(****************************************************************************************************<br>
© Syntegon Group.<br>
All rights reserved, also regarding any disposal, exploitation, reproduction, editing, distribution,<br>
as well as in the event of applications for industrial property rights.<br>
*****************************************************************************************************<br>
DESCRIPTION:<br>
Housekeeping: drops invalid entries and products that have travelled beyond vi_lr_BeltX (along the<br>
conveyor from its start). Products a robot is working on (ASSIGNED or PICKED) are kept wherever they are.<br>
The entries that stay move up in runs (usually one: the products leaving are the oldest, at the front).<br>
*****************************************************************************************************<br>
OUTPUT VALUES:<br>
Number of removed entries.<br>
****************************************************************************************************)
METHOD m_RemoveProductsBeyond : UINT
VAR_INPUT
	vi_lr_BeltX							: LREAL;	// [mm] e.g. belt length + some margin so missed products stay visible briefly
END_VAR
VAR
	un_TempCount						: UINT;	// [-] entries before
	un_TempRead							: UINT;
	un_TempWrite						: UINT;
	un_TempRunStart						: UINT;	// [-] first entry of a run of entries that stay
	b_TempStays							: BOOL;
END_VAR
m_RemoveProductsBeyond := 0;
un_TempCount := vo_Visu.stState.nProductCount;
IF un_TempCount = 0 THEN
	RETURN;
END_IF

(* Keep the entries that stay, in order, moving each run of them up in one go. *)
un_TempWrite := 0;
un_TempRead := 0;
WHILE un_TempRead < un_TempCount DO
	IF m_StaysInRegister(un_TempRead, vi_lr_BeltX) THEN
		un_TempRunStart := un_TempRead;
		b_TempStays := TRUE;
		WHILE b_TempStays DO
			un_TempRead := un_TempRead + 1;
			b_TempStays := FALSE;
			IF un_TempRead < un_TempCount THEN
				b_TempStays := m_StaysInRegister(un_TempRead, vi_lr_BeltX);
			END_IF
		END_WHILE
		IF un_TempWrite <> un_TempRunStart THEN
			Tc2_System.MEMMOVE(ADR(vo_Visu.stState.aProducts[un_TempWrite]), ADR(vo_Visu.stState.aProducts[un_TempRunStart]),
				UINT_TO_UDINT(un_TempRead - un_TempRunStart) * SIZEOF(ST_VisuProduct));
		END_IF
		un_TempWrite := un_TempWrite + (un_TempRead - un_TempRunStart);
	ELSE
		un_TempRead := un_TempRead + 1;
	END_IF
END_WHILE

(* Invalidate the freed tail. *)
m_RemoveProductsBeyond := un_TempCount - un_TempWrite;
IF un_TempWrite < un_TempCount THEN
	FOR un_TempRead := un_TempWrite TO un_TempCount - 1 DO
		vo_Visu.stState.aProducts[un_TempRead].bValid := FALSE;
	END_FOR
	vo_Visu.stState.nProductCount := un_TempWrite;
	vo_Visu.stState.nTimestamp := m_DcTime();
	b_IndexValid := FALSE;
END_IF
END_METHOD

(****************************************************************************************************<br>
© Syntegon Group.<br>
All rights reserved, also regarding any disposal, exploitation, reproduction, editing, distribution,<br>
as well as in the event of applications for industrial property rights.<br>
*****************************************************************************************************<br>
DESCRIPTION:<br>
The rotation of the conveyor's pose as a row-major 3x3 matrix, R = Rz(fRz) * Ry(fRy) * Rx(fRx) as the contract<br>
defines it (ST_VisuPose) and the visualisation applies it, for m_BeltToMcs and m_McsToBelt.<br>
****************************************************************************************************)
METHOD PRIVATE m_Rotation : BOOL
VAR_OUTPUT
	vo_lr_Rotation						: ARRAY[0..8] OF LREAL;	// [-] row by row
END_VAR
VAR
	lr_TempCx							: LREAL;
	lr_TempSx							: LREAL;
	lr_TempCy							: LREAL;
	lr_TempSy							: LREAL;
	lr_TempCz							: LREAL;
	lr_TempSz							: LREAL;
END_VAR
lr_TempCx := COS(vo_Visu.stConfig.stPose.fRx * VISU_GlobalConst.VISU_lr_DEG_TO_RAD);
lr_TempSx := SIN(vo_Visu.stConfig.stPose.fRx * VISU_GlobalConst.VISU_lr_DEG_TO_RAD);
lr_TempCy := COS(vo_Visu.stConfig.stPose.fRy * VISU_GlobalConst.VISU_lr_DEG_TO_RAD);
lr_TempSy := SIN(vo_Visu.stConfig.stPose.fRy * VISU_GlobalConst.VISU_lr_DEG_TO_RAD);
lr_TempCz := COS(vo_Visu.stConfig.stPose.fRz * VISU_GlobalConst.VISU_lr_DEG_TO_RAD);
lr_TempSz := SIN(vo_Visu.stConfig.stPose.fRz * VISU_GlobalConst.VISU_lr_DEG_TO_RAD);
vo_lr_Rotation[0] := lr_TempCz * lr_TempCy;
vo_lr_Rotation[1] := lr_TempCz * lr_TempSy * lr_TempSx - lr_TempSz * lr_TempCx;
vo_lr_Rotation[2] := lr_TempCz * lr_TempSy * lr_TempCx + lr_TempSz * lr_TempSx;
vo_lr_Rotation[3] := lr_TempSz * lr_TempCy;
vo_lr_Rotation[4] := lr_TempSz * lr_TempSy * lr_TempSx + lr_TempCz * lr_TempCx;
vo_lr_Rotation[5] := lr_TempSz * lr_TempSy * lr_TempCx - lr_TempCz * lr_TempSx;
vo_lr_Rotation[6] := -lr_TempSy;
vo_lr_Rotation[7] := lr_TempCy * lr_TempSx;
vo_lr_Rotation[8] := lr_TempCy * lr_TempCx;
m_Rotation := TRUE;
END_METHOD

(****************************************************************************************************<br>
© Syntegon Group.<br>
All rights reserved, also regarding any disposal, exploitation, reproduction, editing, distribution,<br>
as well as in the event of applications for industrial property rights.<br>
*****************************************************************************************************<br>
DESCRIPTION:<br>
Sets the belt position: how far the belt surface has travelled, continuous (no modulo).<br>
Call once per cycle; it also stamps the state with the cycle's DC time.<br>
****************************************************************************************************)
METHOD m_SetBeltPosition : BOOL
VAR_INPUT
	vi_lr_Position						: LREAL;	// [mm]
END_VAR
vo_Visu.stState.fBeltPosition := vi_lr_Position;
vo_Visu.stState.nTimestamp := m_DcTime();
m_SetBeltPosition := TRUE;
END_METHOD

(****************************************************************************************************<br>
© Syntegon Group.<br>
All rights reserved, also regarding any disposal, exploitation, reproduction, editing, distribution,<br>
as well as in the event of applications for industrial property rights.<br>
*****************************************************************************************************<br>
DESCRIPTION:<br>
Sets whether the belt is drawn as a body. A conveyor without one (FALSE) shows only its products, zones and<br>
its axis from the origin to the conveying direction arrow. Default TRUE. TRUE if anything changed.<br>
****************************************************************************************************)
METHOD m_SetBodyVisible : BOOL
VAR_INPUT
	vi_b_Visible						: BOOL;	// TRUE = drawn as a body, FALSE = a conveyor without one
END_VAR
VAR
	TempNew								: ST_VisuConveyorConfig;
END_VAR
TempNew := vo_Visu.stConfig;
TempNew.bBody := vi_b_Visible;
m_SetBodyVisible := m_ApplyConfig(TempNew);
END_METHOD

(****************************************************************************************************<br>
© Syntegon Group.<br>
All rights reserved, also regarding any disposal, exploitation, reproduction, editing, distribution,<br>
as well as in the event of applications for industrial property rights.<br>
*****************************************************************************************************<br>
DESCRIPTION:<br>
Sets or clears the fault of the conveyor: drawn red with the message while active. The fault stays until it<br>
is cleared with m_SetFault(vi_b_Active := FALSE, vi_str_Message := ''). TRUE.<br>
****************************************************************************************************)
METHOD m_SetFault : BOOL
VAR_INPUT
	vi_b_Active							: BOOL;	// TRUE: fault active
	vi_str_Message						: STRING(80);	// shown to the operator; empty shows 'Fault'
END_VAR
vo_Visu.stState.stFault.bActive := vi_b_Active;
vo_Visu.stState.stFault.sMessage := vi_str_Message;
m_SetFault := TRUE;
END_METHOD

(****************************************************************************************************<br>
© Syntegon Group.<br>
All rights reserved, also regarding any disposal, exploitation, reproduction, editing, distribution,<br>
as well as in the event of applications for industrial property rights.<br>
*****************************************************************************************************<br>
DESCRIPTION:<br>
Like m_SetBeltPosition, for a modulo axis: unwraps the position so the belt position stays continuous.<br>
Call once per cycle.<br>
*****************************************************************************************************<br>
LIMITS:<br>
The axis must move less than half a modulo period per cycle.<br>
****************************************************************************************************)
METHOD m_SetModuloBeltPosition : BOOL
VAR_INPUT
	vi_lr_ModuloPosition				: LREAL;	// [mm] in [0, vi_lr_ModuloPeriod)
	vi_lr_ModuloPeriod					: LREAL;	// [mm] <= 0 passes vi_lr_ModuloPosition through unchanged
	vi_b_Reset							: BOOL;	// TRUE: restart the belt position at vi_lr_ModuloPosition
END_VAR
VAR
	lr_TempPosition						: LREAL;	// [mm]
	lr_TempDelta						: LREAL;	// [mm]
END_VAR
IF vi_b_Reset OR NOT b_ModuloInitialised OR vi_lr_ModuloPeriod <= 0 THEN
	lr_TempPosition := vi_lr_ModuloPosition;
	b_ModuloInitialised := TRUE;
ELSE
	lr_TempDelta := vi_lr_ModuloPosition - lr_LastModuloPosition;
	IF lr_TempDelta > vi_lr_ModuloPeriod / 2 THEN
		lr_TempDelta := lr_TempDelta - vi_lr_ModuloPeriod;
	ELSIF lr_TempDelta < -vi_lr_ModuloPeriod / 2 THEN
		lr_TempDelta := lr_TempDelta + vi_lr_ModuloPeriod;
	END_IF
	lr_TempPosition := vo_Visu.stState.fBeltPosition + lr_TempDelta;
END_IF
lr_LastModuloPosition := vi_lr_ModuloPosition;
m_SetModuloBeltPosition := m_SetBeltPosition(lr_TempPosition);
END_METHOD

(****************************************************************************************************<br>
© Syntegon Group.<br>
All rights reserved, also regarding any disposal, exploitation, reproduction, editing, distribution,<br>
as well as in the event of applications for industrial property rights.<br>
*****************************************************************************************************<br>
DESCRIPTION:<br>
Moves the conveyor's coordinate system away from the belt start (stPose), in the belt's local frame. Belt<br>
coordinates (zones' start, end and CCS offset) then count from the shifted origin. TRUE if anything changed.<br>
****************************************************************************************************)
METHOD m_SetOriginShift : BOOL
VAR_INPUT
	vi_lr_X								: LREAL;	// [mm] along the conveying direction
	vi_lr_Y								: LREAL;	// [mm] across the belt, 0 = none
	vi_lr_Z								: LREAL;	// [mm] along the belt surface normal, 0 = none
END_VAR
VAR
	TempNew								: ST_VisuConveyorConfig;
END_VAR
TempNew := vo_Visu.stConfig;
TempNew.stOriginShift.fX := vi_lr_X;
TempNew.stOriginShift.fY := vi_lr_Y;
TempNew.stOriginShift.fZ := vi_lr_Z;
m_SetOriginShift := m_ApplyConfig(TempNew);
END_METHOD

(****************************************************************************************************<br>
© Syntegon Group.<br>
All rights reserved, also regarding any disposal, exploitation, reproduction, editing, distribution,<br>
as well as in the event of applications for industrial property rights.<br>
*****************************************************************************************************<br>
DESCRIPTION:<br>
Marks a product of the register to single it out, e.g. as a sample: the visualisation draws it in the mark's<br>
colour instead of its state colour. 0 removes the mark. The mark stays through m_SetProductState and<br>
m_MoveProduct; a product latched again (e.g. put down on another conveyor) enters unmarked, so mark it there<br>
again. Name the marks once with _FC_VisuSetMarkName.<br>
*****************************************************************************************************<br>
OUTPUT VALUES:<br>
FALSE if the product is not in the register or vi_un_Mark is above VISU_un_MAX_MARKS.<br>
****************************************************************************************************)
METHOD m_SetProductMark : BOOL
VAR_INPUT
	vi_udn_Id							: UDINT;	// [-] product id
	vi_un_Mark							: UINT;	// [-] product mark 1..VISU_un_MAX_MARKS, 0 = none
END_VAR
VAR
	n_TempIndex							: INT;
END_VAR
m_SetProductMark := FALSE;
IF vi_un_Mark > VISU_GlobalConst.VISU_un_MAX_MARKS THEN
	RETURN;
END_IF
n_TempIndex := m_FindProduct(vi_udn_Id);
IF n_TempIndex < 0 THEN
	RETURN;
END_IF
IF vo_Visu.stState.aProducts[n_TempIndex].nMark <> vi_un_Mark THEN
	vo_Visu.stState.aProducts[n_TempIndex].nMark := vi_un_Mark;
	vo_Visu.stState.nTimestamp := m_DcTime();
END_IF
m_SetProductMark := TRUE;
END_METHOD

(****************************************************************************************************<br>
© Syntegon Group.<br>
All rights reserved, also regarding any disposal, exploitation, reproduction, editing, distribution,<br>
as well as in the event of applications for industrial property rights.<br>
*****************************************************************************************************<br>
DESCRIPTION:<br>
Changes a product's state and names the client that changed it: the robot that is assigned to, picks,<br>
places or releases it, the station that rejects it. The state before is kept as ePreviousState when the<br>
state changes; calling it again with the same state keeps it. The product keeps its mark.<br>
FALSE if the product is not in the register.<br>
****************************************************************************************************)
METHOD m_SetProductState : BOOL
VAR_INPUT
	vi_udn_Id							: UDINT;	// [-] product id
	vi_e_State							: E_VisuProductState;
	vi_udn_ClientId						: UDINT;	// [-] manifest id of the client making the change, 0 = none
	vi_udn_MoverId						: UDINT;	// [-] mover of an XTS gantry or loop carrying the product, 0 = none
	vi_udn_FingerId						: UDINT;	// [-] gripper finger (1-based) the product hangs from while picked, 0 = the flange
END_VAR
VAR
	n_TempIndex							: INT;
END_VAR
n_TempIndex := m_FindProduct(vi_udn_Id);
m_SetProductState := n_TempIndex >= 0;
IF m_SetProductState THEN
	IF vo_Visu.stState.aProducts[n_TempIndex].eState <> vi_e_State THEN
		vo_Visu.stState.aProducts[n_TempIndex].ePreviousState := vo_Visu.stState.aProducts[n_TempIndex].eState;
	END_IF
	vo_Visu.stState.aProducts[n_TempIndex].eState := vi_e_State;
	vo_Visu.stState.aProducts[n_TempIndex].nLastClientId := vi_udn_ClientId;
	vo_Visu.stState.aProducts[n_TempIndex].nMoverId := vi_udn_MoverId;
	vo_Visu.stState.aProducts[n_TempIndex].nFingerId := vi_udn_FingerId;
	vo_Visu.stState.nTimestamp := m_DcTime();
END_IF
END_METHOD

(****************************************************************************************************<br>
© Syntegon Group.<br>
All rights reserved, also regarding any disposal, exploitation, reproduction, editing, distribution,<br>
as well as in the event of applications for industrial property rights.<br>
*****************************************************************************************************<br>
DESCRIPTION:<br>
Adds a product type, or updates the one with the same id. FALSE for vi_udn_Id = 0 or a full list. A CYLINDER's<br>
length and width are its diameters (equal: round, different: oval).<br>
****************************************************************************************************)
METHOD m_SetProductType : BOOL
VAR_INPUT
	vi_udn_Id							: UDINT;	// [-] referenced by m_LatchProduct's vi_udn_ProductType
	vi_lr_Length						: LREAL;	// [mm] along the conveying direction
	vi_lr_Width							: LREAL;	// [mm]
	vi_lr_Height						: LREAL;	// [mm]
	vi_e_Shape							: E_VisuProductShape;	// [-] solid of the product, BOX for a plain box
	vi_lr_CornerRadius					: LREAL;	// [mm] rounded vertical edges of a ROUNDED_BOX, 0 for other shapes
END_VAR
VAR
	TempNew								: ST_VisuConveyorConfig;
	un_TempIndex						: UINT;
END_VAR
m_SetProductType := FALSE;
IF vi_udn_Id = 0 THEN
	RETURN;
END_IF
TempNew := vo_Visu.stConfig;
un_TempIndex := 0;
(* ST evaluates both operands of AND: test the index before reading the array. *)
WHILE un_TempIndex < TempNew.nProductTypeCount DO
	IF TempNew.aProductTypes[un_TempIndex].nId = vi_udn_Id THEN
		EXIT;
	END_IF
	un_TempIndex := un_TempIndex + 1;
END_WHILE
IF un_TempIndex >= VISU_GlobalConst_Param.VISU_un_MAX_PRODUCT_TYPES THEN
	RETURN;
END_IF
IF un_TempIndex = TempNew.nProductTypeCount THEN
	TempNew.nProductTypeCount := TempNew.nProductTypeCount + 1;
END_IF
TempNew.aProductTypes[un_TempIndex].nId := vi_udn_Id;
TempNew.aProductTypes[un_TempIndex].fLength := vi_lr_Length;
TempNew.aProductTypes[un_TempIndex].fWidth := vi_lr_Width;
TempNew.aProductTypes[un_TempIndex].fHeight := vi_lr_Height;
TempNew.aProductTypes[un_TempIndex].eShape := vi_e_Shape;
TempNew.aProductTypes[un_TempIndex].fCornerRadius := vi_lr_CornerRadius;
m_ApplyConfig(TempNew);
m_SetProductType := TRUE;
END_METHOD

(****************************************************************************************************<br>
© Syntegon Group.<br>
All rights reserved, also regarding any disposal, exploitation, reproduction, editing, distribution,<br>
as well as in the event of applications for industrial property rights.<br>
*****************************************************************************************************<br>
DESCRIPTION:<br>
Whether register entry vi_un_Index stays in the register for m_RemoveProductsBeyond: it is valid and has not<br>
travelled beyond vi_lr_BeltX, or a robot is working on it (ASSIGNED or PICKED).<br>
****************************************************************************************************)
METHOD PRIVATE m_StaysInRegister : BOOL
VAR_INPUT
	vi_un_Index							: UINT;	// [-] register index
	vi_lr_BeltX							: LREAL;	// [mm] along the conveyor from its start
END_VAR
(* Belt X from the belt start: the latch pose counts from the origin shift and moves with the belt travel. *)
m_StaysInRegister := vo_Visu.stState.aProducts[vi_un_Index].bValid
	AND (vo_Visu.stConfig.stOriginShift.fX + vo_Visu.stState.aProducts[vi_un_Index].stLatchPose.fX
			+ vo_Visu.stState.fBeltPosition - vo_Visu.stState.aProducts[vi_un_Index].fLatchBeltPosition <= vi_lr_BeltX
		OR vo_Visu.stState.aProducts[vi_un_Index].eState = E_VisuProductState.ASSIGNED
		OR vo_Visu.stState.aProducts[vi_un_Index].eState = E_VisuProductState.PICKED);
END_METHOD

END_FUNCTION_BLOCK

// POUs/_FB_VisuComponent
(****************************************************************************************************<br>
© Syntegon Group.<br>
All rights reserved, also regarding any disposal, exploitation, reproduction, editing, distribution,<br>
as well as in the event of applications for industrial property rights.<br>
*****************************************************************************************************<br>
DESCRIPTION:<br>
Base of every visualised component (_FB_VisuConveyor, _FB_VisuDelta, ...). Handles the manifest entry,<br>
the config version and the DC timestamps. Not used directly.<br>
*****************************************************************************************************<br>
VERSION         ¦ DATE       ¦ NAME      ¦ CHANGE<br>
Syn_Visu 3.0.0  ¦ 2026-10-31 ¦ J.Willner ¦ Naming and layout after the TCAT programming guideline<br>
Syn_Visu 8.0.0  ¦ 2026-11-05 ¦ J.Willner ¦ m_Register without vi_str_Path: the symbol path comes from the instance path<br>
Syn_Visu 10.0.0 ¦ 2026-11-14 ¦ J.Willner ¦ m_SetPose for every component; symbol path from _FC_VisuSymbolPath<br>
****************************************************************************************************)
{attribute 'reflection'}
FUNCTION_BLOCK ABSTRACT _FB_VisuComponent
VAR
	RefManifest							: REFERENCE TO ST_VisuManifest;	// set by m_Register
	udn_ComponentId						: UDINT;	// [-] manifest id, 0 = not registered
	(* Device tree path of this instance, e.g. 'RPP_Visu.Syn_Visu_Demo.MAIN.fb_Infeed', set by TwinCAT at initialisation. *)
	{attribute 'instance-path'}
	{attribute 'noinit'}
	str_InstancePath					: STRING(255);
	str_SymbolPath						: STRING(255);	// symbol path of vo_Visu for the manifest, from str_InstancePath on the first m_Register
END_VAR

(****************************************************************************************************<br>
© Syntegon Group.<br>
All rights reserved, also regarding any disposal, exploitation, reproduction, editing, distribution,<br>
as well as in the event of applications for industrial property rights.<br>
*****************************************************************************************************<br>
DESCRIPTION:<br>
Manifest type of the component. Overridden by every derived FB.<br>
****************************************************************************************************)
METHOD PROTECTED m_ComponentType : E_VisuComponentType
m_ComponentType := E_VisuComponentType.NONE;
END_METHOD

(****************************************************************************************************<br>
© Syntegon Group.<br>
All rights reserved, also regarding any disposal, exploitation, reproduction, editing, distribution,<br>
as well as in the event of applications for industrial property rights.<br>
*****************************************************************************************************<br>
DESCRIPTION:<br>
Distributed-clock time of the calling task's current cycle in ns since 2000-01-01; 0 if unknown.<br>
****************************************************************************************************)
METHOD PROTECTED m_DcTime : ULINT
VAR
	dn_TempTaskIndex					: DINT;
END_VAR
dn_TempTaskIndex := Tc2_System.GETCURTASKINDEXEX();
IF dn_TempTaskIndex > 0 THEN
	m_DcTime := LINT_TO_ULINT(TwinCAT_SystemInfoVarList._TaskInfo[dn_TempTaskIndex].DcTaskTime);
ELSE
	m_DcTime := 0;
END_IF
END_METHOD

(****************************************************************************************************<br>
© Syntegon Group.<br>
All rights reserved, also regarding any disposal, exploitation, reproduction, editing, distribution,<br>
as well as in the event of applications for industrial property rights.<br>
*****************************************************************************************************<br>
DESCRIPTION:<br>
Manifest id given to m_Register; 0 while not registered.<br>
****************************************************************************************************)
METHOD m_Id : UDINT
m_Id := udn_ComponentId;
END_METHOD

(****************************************************************************************************<br>
© Syntegon Group.<br>
All rights reserved, also regarding any disposal, exploitation, reproduction, editing, distribution,<br>
as well as in the event of applications for industrial property rights.<br>
*****************************************************************************************************<br>
DESCRIPTION:<br>
Increments the manifest's nConfigVersion so the gateway re-reads the config. No effect before m_Register.<br>
****************************************************************************************************)
METHOD PROTECTED m_NotifyConfigChanged : BOOL
m_NotifyConfigChanged := __ISVALIDREF(RefManifest);
IF m_NotifyConfigChanged THEN
	RefManifest.nConfigVersion := RefManifest.nConfigVersion + 1;
END_IF
END_METHOD

(****************************************************************************************************<br>
© Syntegon Group.<br>
All rights reserved, also regarding any disposal, exploitation, reproduction, editing, distribution,<br>
as well as in the event of applications for industrial property rights.<br>
*****************************************************************************************************<br>
DESCRIPTION:<br>
Where the derived FB keeps its pose in its contract structure, for m_SetPose.<br>
****************************************************************************************************)
METHOD PROTECTED ABSTRACT m_Pose : BOOL
VAR_OUTPUT
	vo_p_Pose							: POINTER TO ST_VisuPose;
END_VAR
END_METHOD

(****************************************************************************************************<br>
© Syntegon Group.<br>
All rights reserved, also regarding any disposal, exploitation, reproduction, editing, distribution,<br>
as well as in the event of applications for industrial property rights.<br>
*****************************************************************************************************<br>
DESCRIPTION:<br>
Adds this component to the manifest; increments nConfigVersion when the entry is new.<br>
Idempotent: call it every cycle, which also keeps the manifest reference valid after an online change.<br>
The symbol path the gateway reads comes from the instance's own path (see _FC_VisuSymbolPath and<br>
VISU_un_INSTANCE_PATH_SKIP).<br>
*****************************************************************************************************<br>
OUTPUT VALUES:<br>
FALSE for vi_udn_Id = 0, an id already used by a different entry, or a full manifest.<br>
****************************************************************************************************)
METHOD m_Register : BOOL
VAR_IN_OUT
	vio_Manifest						: ST_VisuManifest;	// GVL_Visu.stManifest of the application
END_VAR
VAR_INPUT
	vi_udn_Id							: UDINT;	// [-] unique, > 0
	vi_str_Name							: STRING(80);	// display name
END_VAR
VAR
	e_TempType							: E_VisuComponentType;
	un_TempIndex						: UINT;
END_VAR
m_Register := FALSE;
RefManifest REF= vio_Manifest;
(* Always report the contract version of the library actually running, also after an online change. *)
vio_Manifest.nProtocolVersion := VISU_GlobalConst.VISU_un_PROTOCOL_VERSION;
vio_Manifest.sLibraryVersion := VISU_GlobalConst.VISU_str_LIBRARY_VERSION;
e_TempType := m_ComponentType();
IF vi_udn_Id = 0 OR e_TempType = E_VisuComponentType.NONE THEN
	RETURN;
END_IF
IF str_SymbolPath = '' THEN
	str_SymbolPath := _FC_VisuSymbolPath(vio_str_InstancePath := str_InstancePath, vi_str_Member := '.vo_Visu');
END_IF

(* An existing entry with the same id must match exactly. *)
un_TempIndex := 0;
WHILE un_TempIndex < vio_Manifest.nCount AND un_TempIndex < VISU_GlobalConst_Param.VISU_un_MAX_MANIFEST_ENTRIES DO
	IF vio_Manifest.aEntries[un_TempIndex].nId = vi_udn_Id THEN
		m_Register := vio_Manifest.aEntries[un_TempIndex].eType = e_TempType
					AND vio_Manifest.aEntries[un_TempIndex].sName = vi_str_Name
					AND vio_Manifest.aEntries[un_TempIndex].sPath = str_SymbolPath;
		IF m_Register THEN
			udn_ComponentId := vi_udn_Id;
		END_IF
		RETURN;
	END_IF
	un_TempIndex := un_TempIndex + 1;
END_WHILE

(* New entry. *)
IF vio_Manifest.nCount >= VISU_GlobalConst_Param.VISU_un_MAX_MANIFEST_ENTRIES THEN
	RETURN;
END_IF
vio_Manifest.aEntries[vio_Manifest.nCount].nId := vi_udn_Id;
vio_Manifest.aEntries[vio_Manifest.nCount].eType := e_TempType;
vio_Manifest.aEntries[vio_Manifest.nCount].sName := vi_str_Name;
vio_Manifest.aEntries[vio_Manifest.nCount].sPath := str_SymbolPath;
vio_Manifest.nCount := vio_Manifest.nCount + 1;
vio_Manifest.nConfigVersion := vio_Manifest.nConfigVersion + 1;
udn_ComponentId := vi_udn_Id;
m_Register := TRUE;
END_METHOD

(****************************************************************************************************<br>
© Syntegon Group.<br>
All rights reserved, also regarding any disposal, exploitation, reproduction, editing, distribution,<br>
as well as in the event of applications for industrial property rights.<br>
*****************************************************************************************************<br>
DESCRIPTION:<br>
Sets the component's pose in the MCS; where it lies on the component (a conveyor's belt start, a Delta's base<br>
centre, ...) says the guide. A parameter FB of Syn_Config sets it with m_PassOn; m_Configure holds only the<br>
hardware. Increments the config version only when the pose changes, so it may be called every cycle.<br>
*****************************************************************************************************<br>
OUTPUT VALUES:<br>
TRUE if the pose changed.<br>
****************************************************************************************************)
METHOD m_SetPose : BOOL
VAR_INPUT
	vi_Pose								: ST_VisuPose;	// MCS
END_VAR
VAR
	p_TempPose							: POINTER TO ST_VisuPose;
END_VAR
m_SetPose := FALSE;
m_Pose(vo_p_Pose => p_TempPose);
IF p_TempPose = 0 THEN
	RETURN;
END_IF
(* ST_VisuPose holds LREALs only, so a memory compare sees no padding. *)
m_SetPose := Tc2_System.MEMCMP(ADR(vi_Pose), p_TempPose, SIZEOF(vi_Pose)) <> 0;
IF m_SetPose THEN
	p_TempPose^ := vi_Pose;
	m_NotifyConfigChanged();
END_IF
END_METHOD

END_FUNCTION_BLOCK

// POUs/_FB_VisuDelta
(****************************************************************************************************<br>
© Syntegon Group.<br>
All rights reserved, also regarding any disposal, exploitation, reproduction, editing, distribution,<br>
as well as in the event of applications for industrial property rights.<br>
*****************************************************************************************************<br>
DESCRIPTION:<br>
One visualised Delta robot. Typical cycle:<br>
  fb_Delta.m_Register(vio_Manifest := GVL_Visu.stManifest, vi_udn_Id := 10, vi_str_Name := 'Delta 1');<br>
  fb_Delta.m_SetPose(vi_Pose := BasePose);<br>
  fb_Delta.m_Configure(vi_lr_BaseRadius := 200, vi_lr_EffectorRadius := 50,<br>
      vi_lr_UpperArmLength := 400, vi_lr_LowerArmLength := 1000);<br>
  fb_Delta.m_SetFinger(vi_un_Finger := 1, vi_lr_Diameter := 40, vi_lr_Height := 50);<br>
  fb_Delta.m_SetWorkingArea(vi_lr_Radius := 750, vi_lr_ZMin := -1300, vi_lr_ZMax := -700, vi_lr_ConeHeight := 200,<br>
      vi_lr_ConeBottomRadius := 450);<br>
  fb_Delta.m_SetLimitArea(vi_lr_XMin := -500, vi_lr_XMax := 500, vi_lr_YMin := -750, vi_lr_YMax := 750,<br>
      vi_lr_ZMin := -1500, vi_lr_ZMax := -700);<br>
  fb_Delta.m_SetZone(vi_un_Zone := 1, vi_udn_ConveyorId := 1, vi_lr_Start := 1100, vi_lr_End := 1900,<br>
      vi_lr_AllocationOffset := 300, vi_lr_CcsOffset := 1100, vi_lr_StartY := 0, vi_lr_EndY := 0);<br>
  fb_Delta.m_SetTcp(vi_ActualTcp := ActualTcp, vi_SetpointTcp := SetpointTcp);<br>
  fb_Delta.m_SetFingerState(vi_un_Finger := 1, vi_Pose := CupPose, vi_b_Active := b_Vacuum);<br>
Only the TCP (the gripper flange) is reported; the visualisation derives the arms from it. Tool rotations<br>
(e.g. a 4th axis) show only through the finger poses, absolute in the MCS. The config methods may be called<br>
every cycle; the config version only changes when a value does.<br>
*****************************************************************************************************<br>
OUTPUT VALUES:<br>
vo_Visu is the contract structure the gateway reads at the path given to m_Register. Do not write it.<br>
*****************************************************************************************************<br>
VERSION         ¦ DATE       ¦ NAME      ¦ CHANGE<br>
Syn_Visu 3.0.0  ¦ 2026-10-31 ¦ J.Willner ¦ Naming and layout after the TCAT programming guideline<br>
Syn_Visu 4.0.0  ¦ 2026-11-01 ¦ J.Willner ¦ Zones and fingers from _FB_VisuRobot; m_SetZone by index, no kind<br>
Syn_Visu 10.0.0 ¦ 2026-11-14 ¦ J.Willner ¦ Pose by m_SetPose, not m_Configure<br>
****************************************************************************************************)
FUNCTION_BLOCK _FB_VisuDelta EXTENDS _FB_VisuRobot
VAR_OUTPUT
	vo_Visu								: ST_VisuDelta;	// contract structure read by the gateway
END_VAR

(****************************************************************************************************<br>
© Syntegon Group.<br>
All rights reserved, also regarding any disposal, exploitation, reproduction, editing, distribution,<br>
as well as in the event of applications for industrial property rights.<br>
*****************************************************************************************************<br>
DESCRIPTION:<br>
Takes over vio_New and increments the config version if it differs from the current config. TRUE if changed.<br>
****************************************************************************************************)
METHOD PRIVATE m_ApplyConfig : BOOL
VAR_IN_OUT
	vio_New								: ST_VisuDeltaConfig;
END_VAR
m_ApplyConfig := Tc2_System.MEMCMP(ADR(vio_New), ADR(vo_Visu.stConfig), SIZEOF(vio_New)) <> 0;
IF m_ApplyConfig THEN
	vo_Visu.stConfig := vio_New;
	m_NotifyConfigChanged();
END_IF
END_METHOD

(****************************************************************************************************<br>
© Syntegon Group.<br>
All rights reserved, also regarding any disposal, exploitation, reproduction, editing, distribution,<br>
as well as in the event of applications for industrial property rights.<br>
*****************************************************************************************************<br>
DESCRIPTION:<br>
Base pose last set by m_SetPose, MCS.<br>
****************************************************************************************************)
METHOD m_BasePose : ST_VisuPose
m_BasePose := vo_Visu.stConfig.stPose;
END_METHOD

(****************************************************************************************************<br>
© Syntegon Group.<br>
All rights reserved, also regarding any disposal, exploitation, reproduction, editing, distribution,<br>
as well as in the event of applications for industrial property rights.<br>
*****************************************************************************************************<br>
DESCRIPTION:<br>
Manifest type: Delta robot.<br>
****************************************************************************************************)
METHOD PROTECTED m_ComponentType : E_VisuComponentType
m_ComponentType := E_VisuComponentType.DELTA;
END_METHOD

(****************************************************************************************************<br>
© Syntegon Group.<br>
All rights reserved, also regarding any disposal, exploitation, reproduction, editing, distribution,<br>
as well as in the event of applications for industrial property rights.<br>
*****************************************************************************************************<br>
DESCRIPTION:<br>
Sets the geometry; its pose (m_SetPose) is the base centre. Arm 1 lies along the base's local +X; arms 2 and 3 follow<br>
counter-clockwise (seen from above) at 120 deg each. TRUE if anything changed.<br>
****************************************************************************************************)
METHOD m_Configure : BOOL
VAR_INPUT
	vi_lr_BaseRadius					: LREAL;	// [mm] base centre to shoulder joint
	vi_lr_EffectorRadius				: LREAL;	// [mm] effector centre to lower-arm joint
	vi_lr_UpperArmLength				: LREAL;	// [mm]
	vi_lr_LowerArmLength				: LREAL;	// [mm]
END_VAR
VAR
	TempNew								: ST_VisuDeltaConfig;
END_VAR
TempNew := vo_Visu.stConfig;
TempNew.fBaseRadius := vi_lr_BaseRadius;
TempNew.fEffectorRadius := vi_lr_EffectorRadius;
TempNew.fUpperArmLength := vi_lr_UpperArmLength;
TempNew.fLowerArmLength := vi_lr_LowerArmLength;
m_Configure := m_ApplyConfig(TempNew);
END_METHOD

(****************************************************************************************************<br>
© Syntegon Group.<br>
All rights reserved, also regarding any disposal, exploitation, reproduction, editing, distribution,<br>
as well as in the event of applications for industrial property rights.<br>
*****************************************************************************************************<br>
DESCRIPTION:<br>
The robot's gripper fingers for _FB_VisuRobot.m_SetFinger and m_ClearFingers.<br>
****************************************************************************************************)
METHOD PROTECTED m_Fingers : BOOL
VAR_OUTPUT
	vo_p_Count							: POINTER TO UINT;
	vo_p_Fingers						: POINTER TO ARRAY[0..VISU_GlobalConst_Param.VISU_un_MAX_FINGERS - 1] OF ST_VisuFinger;
END_VAR
vo_p_Count := ADR(vo_Visu.stConfig.nFingerCount);
vo_p_Fingers := ADR(vo_Visu.stConfig.aFingers);
m_Fingers := TRUE;
END_METHOD

(****************************************************************************************************<br>
© Syntegon Group.<br>
All rights reserved, also regarding any disposal, exploitation, reproduction, editing, distribution,<br>
as well as in the event of applications for industrial property rights.<br>
*****************************************************************************************************<br>
DESCRIPTION:<br>
The robot's limit area and TCP limit area for _FB_VisuRobot.m_SetLimitArea, m_ClearLimitArea,<br>
m_SetTcpLimitArea and m_ClearTcpLimitArea.<br>
****************************************************************************************************)
METHOD PROTECTED m_LimitArea : BOOL
VAR_OUTPUT
	vo_p_LimitArea						: POINTER TO ST_VisuLimitArea;
	vo_p_TcpLimitArea					: POINTER TO ST_VisuLimitArea;
END_VAR
vo_p_LimitArea := ADR(vo_Visu.stConfig.stLimitArea);
vo_p_TcpLimitArea := ADR(vo_Visu.stConfig.stTcpLimitArea);
m_LimitArea := TRUE;
END_METHOD

(****************************************************************************************************<br>
© Syntegon Group.<br>
All rights reserved, also regarding any disposal, exploitation, reproduction, editing, distribution,<br>
as well as in the event of applications for industrial property rights.<br>
*****************************************************************************************************<br>
DESCRIPTION:<br>
The pose in vo_Visu, for m_SetPose.<br>
****************************************************************************************************)
METHOD PROTECTED m_Pose : BOOL
VAR_OUTPUT
	vo_p_Pose							: POINTER TO ST_VisuPose;
END_VAR
vo_p_Pose := ADR(vo_Visu.stConfig.stPose);
m_Pose := TRUE;
END_METHOD

(****************************************************************************************************<br>
© Syntegon Group.<br>
All rights reserved, also regarding any disposal, exploitation, reproduction, editing, distribution,<br>
as well as in the event of applications for industrial property rights.<br>
*****************************************************************************************************<br>
DESCRIPTION:<br>
Sets or clears the fault of the robot: drawn red with the message while active. The fault stays until it<br>
is cleared with m_SetFault(vi_b_Active := FALSE, vi_str_Message := ''). TRUE.<br>
****************************************************************************************************)
METHOD m_SetFault : BOOL
VAR_INPUT
	vi_b_Active							: BOOL;	// TRUE: fault active
	vi_str_Message						: STRING(80);	// shown to the operator; empty shows 'Fault'
END_VAR
vo_Visu.stState.stFault.bActive := vi_b_Active;
vo_Visu.stState.stFault.sMessage := vi_str_Message;
m_SetFault := TRUE;
END_METHOD

(****************************************************************************************************<br>
© Syntegon Group.<br>
All rights reserved, also regarding any disposal, exploitation, reproduction, editing, distribution,<br>
as well as in the event of applications for industrial property rights.<br>
*****************************************************************************************************<br>
DESCRIPTION:<br>
Reports finger vi_un_Finger (1-based): the pose of its frame (centre of its top face), absolute in the MCS,<br>
and whether it grips. Call once per cycle per configured finger. A finger never reported here is drawn at its<br>
offset on the flange (m_SetFingerOffset, ADR 0018).<br>
*****************************************************************************************************<br>
OUTPUT VALUES:<br>
FALSE outside 1..VISU_GlobalConst_Param.VISU_un_MAX_FINGERS.<br>
****************************************************************************************************)
METHOD m_SetFingerState : BOOL
VAR_INPUT
	vi_un_Finger						: UINT;	// [-] 1-based
	vi_Pose								: ST_VisuPose;	// MCS
	vi_b_Active							: BOOL;	// TRUE while the finger grips
END_VAR
m_SetFingerState := vi_un_Finger > 0 AND vi_un_Finger <= VISU_GlobalConst_Param.VISU_un_MAX_FINGERS;
IF m_SetFingerState THEN
	vo_Visu.stState.aFingerStates[vi_un_Finger - 1].stPose := vi_Pose;
	vo_Visu.stState.aFingerStates[vi_un_Finger - 1].bActive := vi_b_Active;
	vo_Visu.stState.aFingerStates[vi_un_Finger - 1].bPoseReported := TRUE;
END_IF
END_METHOD

(****************************************************************************************************<br>
© Syntegon Group.<br>
All rights reserved, also regarding any disposal, exploitation, reproduction, editing, distribution,<br>
as well as in the event of applications for industrial property rights.<br>
*****************************************************************************************************<br>
DESCRIPTION:<br>
Moves the robot's shown coordinate system (origin triad, local measuring coordinates) away from the base<br>
centre (stPose), in the base's local frame. Geometry, working area and limit area stay relative to stPose.<br>
TRUE if anything changed.<br>
****************************************************************************************************)
METHOD m_SetOriginShift : BOOL
VAR_INPUT
	vi_lr_X								: LREAL;	// [mm] along the base's local X
	vi_lr_Y								: LREAL;	// [mm] along the base's local Y, 0 = none
	vi_lr_Z								: LREAL;	// [mm] along the base's local Z, 0 = none
END_VAR
VAR
	TempNew								: ST_VisuDeltaConfig;
END_VAR
TempNew := vo_Visu.stConfig;
TempNew.stOriginShift.fX := vi_lr_X;
TempNew.stOriginShift.fY := vi_lr_Y;
TempNew.stOriginShift.fZ := vi_lr_Z;
m_SetOriginShift := m_ApplyConfig(TempNew);
END_METHOD

(****************************************************************************************************<br>
© Syntegon Group.<br>
All rights reserved, also regarding any disposal, exploitation, reproduction, editing, distribution,<br>
as well as in the event of applications for industrial property rights.<br>
*****************************************************************************************************<br>
DESCRIPTION:<br>
Reports the robot's TCP. Call once per cycle; it also stamps the state with the cycle's DC time.<br>
****************************************************************************************************)
METHOD m_SetTcp : BOOL
VAR_INPUT
	vi_ActualTcp						: ST_VisuPosition;	// MCS, effector centre (the gripper flange)
	vi_SetpointTcp						: ST_VisuPosition;	// MCS
END_VAR
vo_Visu.stState.stActualTcp := vi_ActualTcp;
vo_Visu.stState.stSetpointTcp := vi_SetpointTcp;
vo_Visu.stState.nTimestamp := m_DcTime();
m_SetTcp := TRUE;
END_METHOD

(****************************************************************************************************<br>
© Syntegon Group.<br>
All rights reserved, also regarding any disposal, exploitation, reproduction, editing, distribution,<br>
as well as in the event of applications for industrial property rights.<br>
*****************************************************************************************************<br>
DESCRIPTION:<br>
Sets the working area: a vertical cylinder in the robot frame with an optional cone below. TRUE if changed.<br>
****************************************************************************************************)
METHOD m_SetWorkingArea : BOOL
VAR_INPUT
	vi_lr_Radius						: LREAL;	// [mm]
	vi_lr_ZMin							: LREAL;	// [mm] relative to the base (below the base: negative)
	vi_lr_ZMax							: LREAL;	// [mm] relative to the base
	vi_lr_ConeHeight					: LREAL;	// [mm] below vi_lr_ZMin; 0 = no cone
	vi_lr_ConeBottomRadius				: LREAL;	// [mm]
END_VAR
VAR
	TempNew								: ST_VisuDeltaConfig;
END_VAR
TempNew := vo_Visu.stConfig;
TempNew.stWorkingArea.fRadius := vi_lr_Radius;
TempNew.stWorkingArea.fZMin := vi_lr_ZMin;
TempNew.stWorkingArea.fZMax := vi_lr_ZMax;
TempNew.stWorkingArea.fConeHeight := vi_lr_ConeHeight;
TempNew.stWorkingArea.fConeBottomRadius := vi_lr_ConeBottomRadius;
m_SetWorkingArea := m_ApplyConfig(TempNew);
END_METHOD

(****************************************************************************************************<br>
© Syntegon Group.<br>
All rights reserved, also regarding any disposal, exploitation, reproduction, editing, distribution,<br>
as well as in the event of applications for industrial property rights.<br>
*****************************************************************************************************<br>
DESCRIPTION:<br>
The robot's zones for _FB_VisuZoneComponent.m_SetZone and m_ClearZones.<br>
****************************************************************************************************)
METHOD PROTECTED m_Zones : BOOL
VAR_OUTPUT
	vo_p_Count							: POINTER TO UINT;
	vo_p_Zones							: POINTER TO ARRAY[0..VISU_GlobalConst_Param.VISU_un_MAX_ZONES - 1] OF ST_VisuZone;
END_VAR
vo_p_Count := ADR(vo_Visu.stConfig.nZoneCount);
vo_p_Zones := ADR(vo_Visu.stConfig.aZones);
m_Zones := TRUE;
END_METHOD

END_FUNCTION_BLOCK

// POUs/_FB_VisuRobot
(****************************************************************************************************<br>
© Syntegon Group.<br>
All rights reserved, also regarding any disposal, exploitation, reproduction, editing, distribution,<br>
as well as in the event of applications for industrial property rights.<br>
*****************************************************************************************************<br>
DESCRIPTION:<br>
Base of every robot (Delta, XTS gantry, XTS loop, Cartesian): zones plus the gripper fingers, m_SetFinger,<br>
m_SetFingerOffset (a finger's place on the flange) and m_ClearFingers, the limit area, m_SetLimitArea and<br>
m_ClearLimitArea, and the TCP limit area, m_SetTcpLimitArea and m_ClearTcpLimitArea. A derived FB tells where<br>
its fingers and its boxes lie through m_Fingers and m_LimitArea; an XTS loop has neither box.<br>
Not used directly.<br>
*****************************************************************************************************<br>
VERSION         ¦ DATE       ¦ NAME      ¦ CHANGE<br>
Syn_Visu 4.0.0  ¦ 2026-11-01 ¦ J.Willner ¦ New: fingers shared by all robots<br>
Syn_Visu 9.3.0  ¦ 2026-11-07 ¦ J.Willner ¦ Limit area shared by Delta, XTS gantry and Cartesian (was Delta only)<br>
Syn_Visu 9.4.0  ¦ 2026-11-09 ¦ J.Willner ¦ TCP limit area: m_SetTcpLimitArea, m_ClearTcpLimitArea<br>
Syn_Visu 9.4.1  ¦ 2026-11-09 ¦ J.Willner ¦ Limit area compares ignore padding: no config change from unchanged values<br>
Syn_Visu 9.5.0  ¦ 2026-11-11 ¦ J.Willner ¦ m_SetFingerOffset: a finger's place on the flange (ADR 0018)<br>
****************************************************************************************************)
FUNCTION_BLOCK ABSTRACT _FB_VisuRobot EXTENDS _FB_VisuZoneComponent

(****************************************************************************************************<br>
© Syntegon Group.<br>
All rights reserved, also regarding any disposal, exploitation, reproduction, editing, distribution,<br>
as well as in the event of applications for industrial property rights.<br>
*****************************************************************************************************<br>
DESCRIPTION:<br>
Removes the gripper definition. TRUE if there was one.<br>
****************************************************************************************************)
METHOD m_ClearFingers : BOOL
VAR
	p_TempCount							: POINTER TO UINT;
	p_TempFingers						: POINTER TO ARRAY[0..VISU_GlobalConst_Param.VISU_un_MAX_FINGERS - 1] OF ST_VisuFinger;
	TempEmpty							: ST_VisuFinger;
	un_TempIndex						: UINT;
END_VAR
m_ClearFingers := FALSE;
m_Fingers(vo_p_Count => p_TempCount, vo_p_Fingers => p_TempFingers);
IF p_TempCount = 0 OR p_TempFingers = 0 THEN
	RETURN;
END_IF
m_ClearFingers := p_TempCount^ > 0;
FOR un_TempIndex := 0 TO VISU_GlobalConst_Param.VISU_un_MAX_FINGERS - 1 DO
	p_TempFingers^[un_TempIndex] := TempEmpty;
END_FOR
p_TempCount^ := 0;
IF m_ClearFingers THEN
	m_NotifyConfigChanged();
END_IF
END_METHOD

(****************************************************************************************************<br>
© Syntegon Group.<br>
All rights reserved, also regarding any disposal, exploitation, reproduction, editing, distribution,<br>
as well as in the event of applications for industrial property rights.<br>
*****************************************************************************************************<br>
DESCRIPTION:<br>
Removes the limit area. TRUE if there was one.<br>
****************************************************************************************************)
METHOD m_ClearLimitArea : BOOL
VAR
	p_TempLimitArea						: POINTER TO ST_VisuLimitArea;
	TempEmpty							: ST_VisuLimitArea;
END_VAR
m_ClearLimitArea := FALSE;
m_LimitArea(vo_p_LimitArea => p_TempLimitArea);
IF p_TempLimitArea = 0 THEN
	RETURN;
END_IF
m_ClearLimitArea := p_TempLimitArea^.bActive;
(* Zeroed first: the MEMCMP below also compares the padding after bActive, which a method local leaves undefined. *)
Tc2_System.MEMSET(ADR(TempEmpty), 0, SIZEOF(TempEmpty));
IF Tc2_System.MEMCMP(ADR(TempEmpty), p_TempLimitArea, SIZEOF(TempEmpty)) <> 0 THEN
	p_TempLimitArea^ := TempEmpty;
	m_NotifyConfigChanged();
END_IF
END_METHOD

(****************************************************************************************************<br>
© Syntegon Group.<br>
All rights reserved, also regarding any disposal, exploitation, reproduction, editing, distribution,<br>
as well as in the event of applications for industrial property rights.<br>
*****************************************************************************************************<br>
DESCRIPTION:<br>
Removes the TCP limit area. TRUE if there was one.<br>
****************************************************************************************************)
METHOD m_ClearTcpLimitArea : BOOL
VAR
	p_TempTcpLimitArea					: POINTER TO ST_VisuLimitArea;
	TempEmpty							: ST_VisuLimitArea;
END_VAR
m_ClearTcpLimitArea := FALSE;
m_LimitArea(vo_p_TcpLimitArea => p_TempTcpLimitArea);
IF p_TempTcpLimitArea = 0 THEN
	RETURN;
END_IF
m_ClearTcpLimitArea := p_TempTcpLimitArea^.bActive;
(* Zeroed first: the MEMCMP below also compares the padding after bActive, which a method local leaves undefined. *)
Tc2_System.MEMSET(ADR(TempEmpty), 0, SIZEOF(TempEmpty));
IF Tc2_System.MEMCMP(ADR(TempEmpty), p_TempTcpLimitArea, SIZEOF(TempEmpty)) <> 0 THEN
	p_TempTcpLimitArea^ := TempEmpty;
	m_NotifyConfigChanged();
END_IF
END_METHOD

(****************************************************************************************************<br>
© Syntegon Group.<br>
All rights reserved, also regarding any disposal, exploitation, reproduction, editing, distribution,<br>
as well as in the event of applications for industrial property rights.<br>
*****************************************************************************************************<br>
DESCRIPTION:<br>
Where the gripper fingers lie in the derived FB's contract structure: vo_p_Count points to its<br>
nFingerCount, vo_p_Fingers to its aFingers.<br>
****************************************************************************************************)
METHOD PROTECTED ABSTRACT m_Fingers : BOOL
VAR_OUTPUT
	vo_p_Count							: POINTER TO UINT;
	vo_p_Fingers						: POINTER TO ARRAY[0..VISU_GlobalConst_Param.VISU_un_MAX_FINGERS - 1] OF ST_VisuFinger;
END_VAR
END_METHOD

(****************************************************************************************************<br>
© Syntegon Group.<br>
All rights reserved, also regarding any disposal, exploitation, reproduction, editing, distribution,<br>
as well as in the event of applications for industrial property rights.<br>
*****************************************************************************************************<br>
DESCRIPTION:<br>
Where the limit area and the TCP limit area lie in the derived FB's contract structure: vo_p_LimitArea points<br>
to its stLimitArea, vo_p_TcpLimitArea to its stTcpLimitArea; both are 0 for a robot without them (XTS loop: it<br>
has no working area of its own).<br>
****************************************************************************************************)
METHOD PROTECTED ABSTRACT m_LimitArea : BOOL
VAR_OUTPUT
	vo_p_LimitArea						: POINTER TO ST_VisuLimitArea;
	vo_p_TcpLimitArea					: POINTER TO ST_VisuLimitArea;
END_VAR
END_METHOD

(****************************************************************************************************<br>
© Syntegon Group.<br>
All rights reserved, also regarding any disposal, exploitation, reproduction, editing, distribution,<br>
as well as in the event of applications for industrial property rights.<br>
*****************************************************************************************************<br>
DESCRIPTION:<br>
Defines gripper finger vi_un_Finger (1-based): a cylinder hanging from the finger's pose along its local -Z.<br>
For XTS kinematics it is a finger of every mover's gripper. The finger count grows to vi_un_Finger.<br>
Its place on the gripper flange comes from m_SetFingerOffset and is kept here.<br>
*****************************************************************************************************<br>
OUTPUT VALUES:<br>
FALSE outside 1..VISU_GlobalConst_Param.VISU_un_MAX_FINGERS.<br>
****************************************************************************************************)
METHOD m_SetFinger : BOOL
VAR_INPUT
	vi_un_Finger						: UINT;	// [-] 1-based, as a product's nFingerId
	vi_lr_Diameter						: LREAL;	// [mm]
	vi_lr_Height						: LREAL;	// [mm] along the finger's local -Z
END_VAR
VAR
	p_TempCount							: POINTER TO UINT;
	p_TempFingers						: POINTER TO ARRAY[0..VISU_GlobalConst_Param.VISU_un_MAX_FINGERS - 1] OF ST_VisuFinger;
	TempFinger							: ST_VisuFinger;
END_VAR
m_SetFinger := FALSE;
IF vi_un_Finger = 0 OR vi_un_Finger > VISU_GlobalConst_Param.VISU_un_MAX_FINGERS THEN
	RETURN;
END_IF
m_Fingers(vo_p_Count => p_TempCount, vo_p_Fingers => p_TempFingers);
IF p_TempCount = 0 OR p_TempFingers = 0 THEN
	RETURN;
END_IF
TempFinger.fDiameter := vi_lr_Diameter;
TempFinger.fHeight := vi_lr_Height;
(* The offset stays as m_SetFingerOffset set it. *)
TempFinger.stOffset := p_TempFingers^[vi_un_Finger - 1].stOffset;
IF vi_un_Finger > p_TempCount^
OR Tc2_System.MEMCMP(ADR(TempFinger), ADR(p_TempFingers^[vi_un_Finger - 1]), SIZEOF(TempFinger)) <> 0
THEN
	p_TempFingers^[vi_un_Finger - 1] := TempFinger;
	p_TempCount^ := MAX(p_TempCount^, vi_un_Finger);
	m_NotifyConfigChanged();
END_IF
m_SetFinger := TRUE;
END_METHOD

(****************************************************************************************************<br>
© Syntegon Group.<br>
All rights reserved, also regarding any disposal, exploitation, reproduction, editing, distribution,<br>
as well as in the event of applications for industrial property rights.<br>
*****************************************************************************************************<br>
DESCRIPTION:<br>
Places finger vi_un_Finger (1-based, defined with m_SetFinger) on the gripper flange (ADR 0018): the position<br>
of its frame in the flange frame and its rotation about the flange's Z. The flange frame's -Z points to the<br>
product: a Delta's lies at the TCP with the robot's axes, a Cartesian robot's has the robot's axes, an XTS mover's<br>
turns with the mover. While the application reports no pose for the finger (m_SetFingerState, or an XTS track<br>
with m_SetFingersOnFlange), the visualisation draws it there. The config version only changes when a value does.<br>
*****************************************************************************************************<br>
OUTPUT VALUES:<br>
FALSE for a finger outside 1..the finger count.<br>
****************************************************************************************************)
METHOD m_SetFingerOffset : BOOL
VAR_INPUT
	vi_un_Finger						: UINT;	// [-] 1-based
	vi_lr_X								: LREAL;	// [mm] along the flange's X
	vi_lr_Y								: LREAL;	// [mm] along the flange's Y
	vi_lr_Z								: LREAL;	// [mm] along the flange's Z (towards the product: negative)
	vi_lr_Rz							: LREAL;	// [deg] about the flange's Z
END_VAR
VAR
	p_TempCount							: POINTER TO UINT;
	p_TempFingers						: POINTER TO ARRAY[0..VISU_GlobalConst_Param.VISU_un_MAX_FINGERS - 1] OF ST_VisuFinger;
	TempOffset							: ST_VisuPlanarPose;
END_VAR
m_SetFingerOffset := FALSE;
m_Fingers(vo_p_Count => p_TempCount, vo_p_Fingers => p_TempFingers);
IF p_TempCount = 0 OR p_TempFingers = 0 THEN
	RETURN;
END_IF
IF vi_un_Finger = 0 OR vi_un_Finger > p_TempCount^ THEN
	RETURN;
END_IF
TempOffset.fX := vi_lr_X;
TempOffset.fY := vi_lr_Y;
TempOffset.fZ := vi_lr_Z;
TempOffset.fRz := vi_lr_Rz;
IF Tc2_System.MEMCMP(ADR(TempOffset), ADR(p_TempFingers^[vi_un_Finger - 1].stOffset), SIZEOF(TempOffset)) <> 0 THEN
	p_TempFingers^[vi_un_Finger - 1].stOffset := TempOffset;
	m_NotifyConfigChanged();
END_IF
m_SetFingerOffset := TRUE;
END_METHOD

(****************************************************************************************************<br>
© Syntegon Group.<br>
All rights reserved, also regarding any disposal, exploitation, reproduction, editing, distribution,<br>
as well as in the event of applications for industrial property rights.<br>
*****************************************************************************************************<br>
DESCRIPTION:<br>
Sets and activates the limit area: an axis-aligned box in the robot frame (relative to its pose, the frame its<br>
working area is given in) that further restricts the working area. Delta, XTS gantry and Cartesian robot;<br>
an XTS loop has none. Equal bounds make a flat box. The config version only changes when a value does.<br>
*****************************************************************************************************<br>
OUTPUT VALUES:<br>
TRUE if anything changed; FALSE for a robot without a limit area (XTS loop).<br>
****************************************************************************************************)
METHOD m_SetLimitArea : BOOL
VAR_INPUT
	vi_lr_XMin							: LREAL;	// [mm] in the robot frame
	vi_lr_XMax							: LREAL;	// [mm]
	vi_lr_YMin							: LREAL;	// [mm]
	vi_lr_YMax							: LREAL;	// [mm]
	vi_lr_ZMin							: LREAL;	// [mm] relative to the pose (below it: negative)
	vi_lr_ZMax							: LREAL;	// [mm]
END_VAR
VAR
	p_TempLimitArea						: POINTER TO ST_VisuLimitArea;
	TempLimitArea						: ST_VisuLimitArea;
END_VAR
m_SetLimitArea := FALSE;
m_LimitArea(vo_p_LimitArea => p_TempLimitArea);
IF p_TempLimitArea = 0 THEN
	RETURN;
END_IF
(* Zeroed first: the MEMCMP below also compares the padding after bActive, which a method local leaves undefined. *)
Tc2_System.MEMSET(ADR(TempLimitArea), 0, SIZEOF(TempLimitArea));
TempLimitArea.fXMin := vi_lr_XMin;
TempLimitArea.fXMax := vi_lr_XMax;
TempLimitArea.fYMin := vi_lr_YMin;
TempLimitArea.fYMax := vi_lr_YMax;
TempLimitArea.fZMin := vi_lr_ZMin;
TempLimitArea.fZMax := vi_lr_ZMax;
TempLimitArea.bActive := TRUE;
IF Tc2_System.MEMCMP(ADR(TempLimitArea), p_TempLimitArea, SIZEOF(TempLimitArea)) <> 0 THEN
	p_TempLimitArea^ := TempLimitArea;
	m_NotifyConfigChanged();
	m_SetLimitArea := TRUE;
END_IF
END_METHOD

(****************************************************************************************************<br>
© Syntegon Group.<br>
All rights reserved, also regarding any disposal, exploitation, reproduction, editing, distribution,<br>
as well as in the event of applications for industrial property rights.<br>
*****************************************************************************************************<br>
DESCRIPTION:<br>
Sets and activates the TCP limit area: an axis-aligned box around the TCP (XTS gantry: around every mover's<br>
gripper flange), its bounds relative to the TCP along the axes of the robot frame. It moves with the TCP and<br>
never turns. The visualisation lights it up red with a message when it overlaps another robot's limit area or<br>
TCP limit area (also another mover's of the same gantry), or leaves the robot's own limit area. Delta, XTS<br>
gantry and Cartesian robot; an XTS loop has none. Equal bounds make a flat box. The config version only<br>
changes when a value does.<br>
*****************************************************************************************************<br>
OUTPUT VALUES:<br>
TRUE if anything changed; FALSE for a robot without a TCP limit area (XTS loop).<br>
****************************************************************************************************)
METHOD m_SetTcpLimitArea : BOOL
VAR_INPUT
	vi_lr_XMin							: LREAL;	// [mm] relative to the TCP, along the robot frame's X
	vi_lr_XMax							: LREAL;	// [mm]
	vi_lr_YMin							: LREAL;	// [mm]
	vi_lr_YMax							: LREAL;	// [mm]
	vi_lr_ZMin							: LREAL;	// [mm] relative to the TCP (below it: negative)
	vi_lr_ZMax							: LREAL;	// [mm]
END_VAR
VAR
	p_TempTcpLimitArea					: POINTER TO ST_VisuLimitArea;
	TempTcpLimitArea					: ST_VisuLimitArea;
END_VAR
m_SetTcpLimitArea := FALSE;
m_LimitArea(vo_p_TcpLimitArea => p_TempTcpLimitArea);
IF p_TempTcpLimitArea = 0 THEN
	RETURN;
END_IF
(* Zeroed first: the MEMCMP below also compares the padding after bActive, which a method local leaves undefined. *)
Tc2_System.MEMSET(ADR(TempTcpLimitArea), 0, SIZEOF(TempTcpLimitArea));
TempTcpLimitArea.fXMin := vi_lr_XMin;
TempTcpLimitArea.fXMax := vi_lr_XMax;
TempTcpLimitArea.fYMin := vi_lr_YMin;
TempTcpLimitArea.fYMax := vi_lr_YMax;
TempTcpLimitArea.fZMin := vi_lr_ZMin;
TempTcpLimitArea.fZMax := vi_lr_ZMax;
TempTcpLimitArea.bActive := TRUE;
IF Tc2_System.MEMCMP(ADR(TempTcpLimitArea), p_TempTcpLimitArea, SIZEOF(TempTcpLimitArea)) <> 0 THEN
	p_TempTcpLimitArea^ := TempTcpLimitArea;
	m_NotifyConfigChanged();
	m_SetTcpLimitArea := TRUE;
END_IF
END_METHOD

END_FUNCTION_BLOCK

// POUs/_FB_VisuZoneComponent
(****************************************************************************************************<br>
© Syntegon Group.<br>
All rights reserved, also regarding any disposal, exploitation, reproduction, editing, distribution,<br>
as well as in the event of applications for industrial property rights.<br>
*****************************************************************************************************<br>
DESCRIPTION:<br>
Base of every component with zones on conveyors (robots, detectors): m_SetZone and m_ClearZones.<br>
A derived FB tells where its zones lie in its contract structure through m_Zones. Not used directly.<br>
*****************************************************************************************************<br>
VERSION         ¦ DATE       ¦ NAME      ¦ CHANGE<br>
Syn_Visu 4.0.0  ¦ 2026-11-01 ¦ J.Willner ¦ New: zones shared by robots and detectors, no zone kind<br>
Syn_Visu 9.0.0  ¦ 2026-11-05 ¦ J.Willner ¦ m_SetZone: vi_lr_StartY, vi_lr_EndY bound the zone across the belt<br>
Syn_Visu 9.4.1  ¦ 2026-11-09 ¦ J.Willner ¦ m_SetZone compare ignores padding: no config change from an unchanged zone<br>
****************************************************************************************************)
FUNCTION_BLOCK ABSTRACT _FB_VisuZoneComponent EXTENDS _FB_VisuComponent

(****************************************************************************************************<br>
© Syntegon Group.<br>
All rights reserved, also regarding any disposal, exploitation, reproduction, editing, distribution,<br>
as well as in the event of applications for industrial property rights.<br>
*****************************************************************************************************<br>
DESCRIPTION:<br>
Removes all zones. TRUE if there were any.<br>
****************************************************************************************************)
METHOD m_ClearZones : BOOL
VAR
	p_TempCount							: POINTER TO UINT;
	p_TempZones							: POINTER TO ARRAY[0..VISU_GlobalConst_Param.VISU_un_MAX_ZONES - 1] OF ST_VisuZone;
	TempEmpty							: ST_VisuZone;
	un_TempIndex						: UINT;
END_VAR
m_ClearZones := FALSE;
m_Zones(vo_p_Count => p_TempCount, vo_p_Zones => p_TempZones);
IF p_TempCount = 0 OR p_TempZones = 0 THEN
	RETURN;
END_IF
m_ClearZones := p_TempCount^ > 0;
FOR un_TempIndex := 0 TO VISU_GlobalConst_Param.VISU_un_MAX_ZONES - 1 DO
	p_TempZones^[un_TempIndex] := TempEmpty;
END_FOR
p_TempCount^ := 0;
IF m_ClearZones THEN
	m_NotifyConfigChanged();
END_IF
END_METHOD

(****************************************************************************************************<br>
© Syntegon Group.<br>
All rights reserved, also regarding any disposal, exploitation, reproduction, editing, distribution,<br>
as well as in the event of applications for industrial property rights.<br>
*****************************************************************************************************<br>
DESCRIPTION:<br>
Sets zone vi_un_Zone (1-based): a stretch of a conveyor that belongs to this component, e.g. where a<br>
robot picks or places or where a detector detects. vi_lr_Start = vi_lr_End is a line across the belt;<br>
vi_lr_StartY = vi_lr_EndY spans the whole belt width, else the zone lies between them across the belt.<br>
The zone count grows to vi_un_Zone; set the zones in order. The config version only changes when a<br>
value does.<br>
*****************************************************************************************************<br>
OUTPUT VALUES:<br>
FALSE for vi_udn_ConveyorId = 0 or vi_un_Zone outside 1..VISU_GlobalConst_Param.VISU_un_MAX_ZONES.<br>
****************************************************************************************************)
METHOD m_SetZone : BOOL
VAR_INPUT
	vi_un_Zone							: UINT;	// [-] 1-based
	vi_udn_ConveyorId					: UDINT;	// [-] manifest id of the conveyor
	vi_lr_Start							: LREAL;	// [mm] along the conveyor from its origin (belt coordinates, not MCS)
	vi_lr_End							: LREAL;	// [mm] along the conveyor from its origin
	vi_lr_AllocationOffset				: LREAL;	// [mm] before vi_lr_End up to which products may be allocated; 0 = no limit
	vi_lr_CcsOffset						: LREAL;	// [mm] along the conveyor from its origin: the component's conveyor coordinate system, 0 = its origin
	vi_lr_StartY						: LREAL;	// [mm] across the conveyor from its origin (local Y): one side of the zone
	vi_lr_EndY							: LREAL;	// [mm] across the conveyor from its origin: the other side; = vi_lr_StartY for the whole belt width
END_VAR
VAR
	p_TempCount							: POINTER TO UINT;
	p_TempZones							: POINTER TO ARRAY[0..VISU_GlobalConst_Param.VISU_un_MAX_ZONES - 1] OF ST_VisuZone;
	TempZone							: ST_VisuZone;
END_VAR
m_SetZone := FALSE;
IF vi_udn_ConveyorId = 0 OR vi_un_Zone = 0 OR vi_un_Zone > VISU_GlobalConst_Param.VISU_un_MAX_ZONES THEN
	RETURN;
END_IF
m_Zones(vo_p_Count => p_TempCount, vo_p_Zones => p_TempZones);
IF p_TempCount = 0 OR p_TempZones = 0 THEN
	RETURN;
END_IF
(* Zeroed first: the MEMCMP below also compares the padding after nConveyorId, which a method local leaves undefined. *)
Tc2_System.MEMSET(ADR(TempZone), 0, SIZEOF(TempZone));
TempZone.nConveyorId := vi_udn_ConveyorId;
TempZone.fStart := vi_lr_Start;
TempZone.fEnd := vi_lr_End;
TempZone.fAllocationOffset := vi_lr_AllocationOffset;
TempZone.fCcsOffset := vi_lr_CcsOffset;
TempZone.fStartY := vi_lr_StartY;
TempZone.fEndY := vi_lr_EndY;
IF vi_un_Zone > p_TempCount^
OR Tc2_System.MEMCMP(ADR(TempZone), ADR(p_TempZones^[vi_un_Zone - 1]), SIZEOF(TempZone)) <> 0
THEN
	p_TempZones^[vi_un_Zone - 1] := TempZone;
	p_TempCount^ := MAX(p_TempCount^, vi_un_Zone);
	m_NotifyConfigChanged();
END_IF
m_SetZone := TRUE;
END_METHOD

(****************************************************************************************************<br>
© Syntegon Group.<br>
All rights reserved, also regarding any disposal, exploitation, reproduction, editing, distribution,<br>
as well as in the event of applications for industrial property rights.<br>
*****************************************************************************************************<br>
DESCRIPTION:<br>
Where the zones lie in the derived FB's contract structure: vo_p_Count points to its nZoneCount,<br>
vo_p_Zones to its aZones.<br>
****************************************************************************************************)
METHOD PROTECTED ABSTRACT m_Zones : BOOL
VAR_OUTPUT
	vo_p_Count							: POINTER TO UINT;
	vo_p_Zones							: POINTER TO ARRAY[0..VISU_GlobalConst_Param.VISU_un_MAX_ZONES - 1] OF ST_VisuZone;
END_VAR
END_METHOD

END_FUNCTION_BLOCK

// POUs/_FC_VisuSymbolPath
(****************************************************************************************************<br>
© Syntegon Group.<br>
All rights reserved, also regarding any disposal, exploitation, reproduction, editing, distribution,<br>
as well as in the event of applications for industrial property rights.<br>
*****************************************************************************************************<br>
DESCRIPTION:<br>
The symbol path the gateway reads over ADS for an FB's contract structure, from the FB's instance path: without<br>
the leading VISU_un_INSTANCE_PATH_SKIP segments (TwinCAT project and PLC project), with vi_str_Member appended.<br>
'RPP_Visu.Syn_Visu_Demo.P_VisuDemoDelta.fb_Infeed1' and '.vo_Visu' give 'P_VisuDemoDelta.fb_Infeed1.vo_Visu'.<br>
An instance path with fewer segments is kept whole. Used by the manifests of Syn_Visu and Syn_Config.<br>
*****************************************************************************************************<br>
OUTPUT VALUES:<br>
The symbol path, cut at 255 bytes.<br>
*****************************************************************************************************<br>
VERSION         ¦ DATE       ¦ NAME      ¦ CHANGE<br>
Syn_Visu 10.0.0 ¦ 2026-11-14 ¦ J.Willner ¦ Created: one rule for both manifests<br>
****************************************************************************************************)
FUNCTION _FC_VisuSymbolPath : STRING(255)
VAR_IN_OUT CONSTANT
	vio_str_InstancePath				: STRING(255);	// the FB's {attribute 'instance-path'} variable
END_VAR
VAR_INPUT
	vi_str_Member						: STRING(15);	// the contract structure, e.g. '.vo_Visu'
END_VAR
VAR
	un_TempRead							: UINT;	// [-] byte index in vio_str_InstancePath
	un_TempWrite						: UINT;	// [-] byte index in the result
	un_TempDots							: UINT;	// [-] dots passed
END_VAR
VAR CONSTANT
	un_MAX_INDEX						: UINT := 255;	// [-] last byte of a STRING(255), its terminating zero
	by_DOT								: BYTE := 16#2E;	// '.'
	un_MAX_MEMBER_INDEX					: UINT := 15;	// [-] last byte of vi_str_Member, a STRING(15)
END_VAR

(* Skip the leading segments, up to and including the VISU_un_INSTANCE_PATH_SKIP-th dot. *)
un_TempRead := 0;
un_TempDots := 0;
WHILE un_TempDots < VISU_GlobalConst_Param.VISU_un_INSTANCE_PATH_SKIP AND un_TempRead < un_MAX_INDEX
	AND vio_str_InstancePath[un_TempRead] <> 0
DO
	IF vio_str_InstancePath[un_TempRead] = by_DOT THEN
		un_TempDots := un_TempDots + 1;
	END_IF
	un_TempRead := un_TempRead + 1;
END_WHILE
IF un_TempDots < VISU_GlobalConst_Param.VISU_un_INSTANCE_PATH_SKIP THEN
	un_TempRead := 0;
END_IF

(* The rest of the instance path, then the contract structure. *)
un_TempWrite := 0;
WHILE un_TempRead < un_MAX_INDEX AND vio_str_InstancePath[un_TempRead] <> 0 AND un_TempWrite < un_MAX_INDEX DO
	_FC_VisuSymbolPath[un_TempWrite] := vio_str_InstancePath[un_TempRead];
	un_TempRead := un_TempRead + 1;
	un_TempWrite := un_TempWrite + 1;
END_WHILE
un_TempRead := 0;
WHILE un_TempRead < un_MAX_MEMBER_INDEX AND vi_str_Member[un_TempRead] <> 0 AND un_TempWrite < un_MAX_INDEX DO
	_FC_VisuSymbolPath[un_TempWrite] := vi_str_Member[un_TempRead];
	un_TempRead := un_TempRead + 1;
	un_TempWrite := un_TempWrite + 1;
END_WHILE
_FC_VisuSymbolPath[un_TempWrite] := 0;

END_FUNCTION

// POUs/_FC_VisuSetMarkName
(****************************************************************************************************<br>
© Syntegon Group.<br>
All rights reserved, also regarding any disposal, exploitation, reproduction, editing, distribution,<br>
as well as in the event of applications for industrial property rights.<br>
*****************************************************************************************************<br>
DESCRIPTION:<br>
Names a product mark for the whole PLC in the manifest, e.g. 1 = 'Sample': the visualisation shows the name<br>
with a marked product (_FB_VisuConveyor.m_SetProductMark). An empty name leaves the mark unnamed. Increments<br>
nConfigVersion only when the name changes, so it may be called every cycle.<br>
*****************************************************************************************************<br>
OUTPUT VALUES:<br>
TRUE if the name changed. FALSE for an unchanged name, vi_un_Mark = 0 or one above VISU_un_MAX_MARKS.<br>
*****************************************************************************************************<br>
VERSION         ¦ DATE       ¦ NAME      ¦ CHANGE<br>
Syn_Visu 9.6.0  ¦ 2026-11-12 ¦ J.Willner ¦ Created: product marks (protocol 21)<br>
****************************************************************************************************)
FUNCTION _FC_VisuSetMarkName : BOOL
VAR_IN_OUT
	vio_Manifest						: ST_VisuManifest;	// GVL_Visu.stManifest of the application
END_VAR
VAR_INPUT
	vi_un_Mark							: UINT;	// [-] product mark 1..VISU_un_MAX_MARKS
	vi_str_Name							: STRING(31);	// what the mark means, '' = unnamed
END_VAR

_FC_VisuSetMarkName := FALSE;
IF vi_un_Mark = 0 OR vi_un_Mark > VISU_GlobalConst.VISU_un_MAX_MARKS THEN
	RETURN;
END_IF
IF vio_Manifest.aMarkNames[vi_un_Mark] <> vi_str_Name THEN
	vio_Manifest.aMarkNames[vi_un_Mark] := vi_str_Name;
	vio_Manifest.nConfigVersion := vio_Manifest.nConfigVersion + 1;
	_FC_VisuSetMarkName := TRUE;
END_IF

END_FUNCTION

// POUs/_FB_VisuStation
(****************************************************************************************************<br>
© Syntegon Group.<br>
All rights reserved, also regarding any disposal, exploitation, reproduction, editing, distribution,<br>
as well as in the event of applications for industrial property rights.<br>
*****************************************************************************************************<br>
DESCRIPTION:<br>
One visualised station: a client at a conveyor that works on the products in its zones, e.g. a reject<br>
unit, a labeller, a printer or a check weigher. It is drawn only from the bodies it describes. Typical cycle<br>
of a reject unit:<br>
  fb_Reject.m_Register(vio_Manifest := GVL_Visu.stManifest, vi_udn_Id := 70, vi_str_Name := 'Reject unit');<br>
  fb_Reject.m_SetPose(vi_Pose := StationPose);<br>
  fb_Reject.m_SetBody(vi_un_Body := 1, ...);   // housing<br>
  fb_Reject.m_SetBody(vi_un_Body := 2, ...);   // pusher<br>
  fb_Reject.m_SetZone(vi_un_Zone := 1, vi_udn_ConveyorId := 2, vi_lr_Start := 2400, vi_lr_End := 2400,<br>
      vi_lr_AllocationOffset := 0, vi_lr_CcsOffset := 2400, vi_lr_StartY := 0, vi_lr_EndY := 0);<br>
  fb_Reject.m_SetBodyActive(vi_un_Body := 2, vi_b_Active := b_Pushing);<br>
and on the conveyor, when it rejects a product:<br>
  fb_Outfeed.m_SetProductState(vi_udn_Id := udn_Product, vi_e_State := E_VisuProductState.REJECTED,<br>
      vi_udn_ClientId := fb_Reject.m_Id(), vi_udn_MoverId := 0, vi_udn_FingerId := 0);<br>
A station may also latch products (m_LatchProduct with vi_udn_ClientId := its id), e.g. a check weigher.<br>
*****************************************************************************************************<br>
OUTPUT VALUES:<br>
vo_Visu is the contract structure the gateway reads at the path given to m_Register. Do not write it.<br>
*****************************************************************************************************<br>
VERSION         ¦ DATE       ¦ NAME      ¦ CHANGE<br>
Syn_Visu 6.0.0  ¦ 2026-11-01 ¦ J.Willner ¦ New<br>
Syn_Visu 10.0.0 ¦ 2026-11-14 ¦ J.Willner ¦ Pose by m_SetPose; m_Configure removed<br>
****************************************************************************************************)
FUNCTION_BLOCK _FB_VisuStation EXTENDS _FB_VisuBodyComponent
VAR_OUTPUT
	vo_Visu								: ST_VisuStation;	// contract structure read by the gateway
END_VAR

(****************************************************************************************************<br>
© Syntegon Group.<br>
All rights reserved, also regarding any disposal, exploitation, reproduction, editing, distribution,<br>
as well as in the event of applications for industrial property rights.<br>
*****************************************************************************************************<br>
DESCRIPTION:<br>
Manifest type: station.<br>
****************************************************************************************************)
METHOD PROTECTED m_ComponentType : E_VisuComponentType
m_ComponentType := E_VisuComponentType.STATION;
END_METHOD

(****************************************************************************************************<br>
© Syntegon Group.<br>
All rights reserved, also regarding any disposal, exploitation, reproduction, editing, distribution,<br>
as well as in the event of applications for industrial property rights.<br>
*****************************************************************************************************<br>
DESCRIPTION:<br>
The station's pose, origin shift, bodies, body states, timestamp and fault for _FB_VisuBodyComponent.<br>
****************************************************************************************************)
METHOD PROTECTED m_Parts : BOOL
VAR_OUTPUT
	vo_p_Pose							: POINTER TO ST_VisuPose;
	vo_p_OriginShift					: POINTER TO ST_VisuPosition;
	vo_p_BodyCount						: POINTER TO UINT;
	vo_p_Bodies							: POINTER TO ARRAY[0..VISU_GlobalConst_Param.VISU_un_MAX_BODIES - 1] OF ST_VisuBody;
	vo_p_BodyStates						: POINTER TO ARRAY[0..VISU_GlobalConst_Param.VISU_un_MAX_BODIES - 1] OF ST_VisuBodyState;
	vo_p_Timestamp						: POINTER TO ULINT;
	vo_p_Fault							: POINTER TO ST_VisuFault;
END_VAR
vo_p_Pose := ADR(vo_Visu.stConfig.stPose);
vo_p_OriginShift := ADR(vo_Visu.stConfig.stOriginShift);
vo_p_BodyCount := ADR(vo_Visu.stConfig.nBodyCount);
vo_p_Bodies := ADR(vo_Visu.stConfig.aBodies);
vo_p_BodyStates := ADR(vo_Visu.stState.aBodyStates);
vo_p_Timestamp := ADR(vo_Visu.stState.nTimestamp);
vo_p_Fault := ADR(vo_Visu.stState.stFault);
m_Parts := TRUE;
END_METHOD

(****************************************************************************************************<br>
© Syntegon Group.<br>
All rights reserved, also regarding any disposal, exploitation, reproduction, editing, distribution,<br>
as well as in the event of applications for industrial property rights.<br>
*****************************************************************************************************<br>
DESCRIPTION:<br>
The station's zones for _FB_VisuZoneComponent.m_SetZone and m_ClearZones.<br>
****************************************************************************************************)
METHOD PROTECTED m_Zones : BOOL
VAR_OUTPUT
	vo_p_Count							: POINTER TO UINT;
	vo_p_Zones							: POINTER TO ARRAY[0..VISU_GlobalConst_Param.VISU_un_MAX_ZONES - 1] OF ST_VisuZone;
END_VAR
vo_p_Count := ADR(vo_Visu.stConfig.nZoneCount);
vo_p_Zones := ADR(vo_Visu.stConfig.aZones);
m_Zones := TRUE;
END_METHOD

END_FUNCTION_BLOCK

// POUs/_FB_VisuCartesian
(****************************************************************************************************<br>
© Syntegon Group.<br>
All rights reserved, also regarding any disposal, exploitation, reproduction, editing, distribution,<br>
as well as in the event of applications for industrial property rights.<br>
*****************************************************************************************************<br>
DESCRIPTION:<br>
One visualised Cartesian robot: linear X, Y, Z axes ending at a gripper flange; m_SetKinematics leaves out the<br>
Y axis (XZ, a fixed beam) or the Z axis (XY). Typical cycle:<br>
  fb_Cartesian.m_Register(vio_Manifest := GVL_Visu.stManifest, vi_udn_Id := 40, vi_str_Name := 'Cartesian');<br>
  fb_Cartesian.m_SetPose(vi_Pose := RobotPose);<br>
  fb_Cartesian.m_Configure(vi_lr_XMin := 0, vi_lr_XMax := 1200, vi_lr_YMin := 0,<br>
      vi_lr_YMax := 1000, vi_lr_ZMin := -600, vi_lr_ZMax := 0, vi_lr_RailHeight := 1200);<br>
  fb_Cartesian.m_SetFinger(vi_un_Finger := 1, vi_lr_Diameter := 40, vi_lr_Height := 40);<br>
  fb_Cartesian.m_SetZone(vi_un_Zone := 1, vi_udn_ConveyorId := 7, vi_lr_Start := 1000, vi_lr_End := 2000,<br>
      vi_lr_AllocationOffset := 0, vi_lr_CcsOffset := 1000, vi_lr_StartY := 0, vi_lr_EndY := 0);<br>
  fb_Cartesian.m_SetAxes(vi_lr_X := ..., vi_lr_Y := ..., vi_lr_Z := ..., vi_b_GripperActive := ...);<br>
  fb_Cartesian.m_SetFingerState(vi_un_Finger := 1, vi_Pose := CupPose, vi_b_Active := b_Vacuum);<br>
Only actual values are reported; tool rotations (e.g. C and A) show only through the finger poses, absolute in<br>
the MCS. The config methods may be called every cycle; the config version only changes when a value does.<br>
*****************************************************************************************************<br>
OUTPUT VALUES:<br>
vo_Visu is the contract structure the gateway reads at the path given to m_Register. Do not write it.<br>
*****************************************************************************************************<br>
VERSION         ¦ DATE       ¦ NAME      ¦ CHANGE<br>
Syn_Visu 3.0.0  ¦ 2026-10-31 ¦ J.Willner ¦ Naming and layout after the TCAT programming guideline<br>
Syn_Visu 4.0.0  ¦ 2026-11-01 ¦ J.Willner ¦ Zones and fingers from _FB_VisuRobot; m_SetZone by index, no kind<br>
Syn_Visu 9.2.0  ¦ 2026-11-07 ¦ J.Willner ¦ m_SetKinematics: without Y axis (XZ) or Z axis (XY)<br>
Syn_Visu 10.0.0 ¦ 2026-11-14 ¦ J.Willner ¦ Pose by m_SetPose, not m_Configure<br>
****************************************************************************************************)
FUNCTION_BLOCK _FB_VisuCartesian EXTENDS _FB_VisuRobot
VAR_OUTPUT
	vo_Visu								: ST_VisuCartesian;	// contract structure read by the gateway
END_VAR

(****************************************************************************************************<br>
© Syntegon Group.<br>
All rights reserved, also regarding any disposal, exploitation, reproduction, editing, distribution,<br>
as well as in the event of applications for industrial property rights.<br>
*****************************************************************************************************<br>
DESCRIPTION:<br>
Takes over vio_New and increments the config version if it differs from the current config. TRUE if changed.<br>
****************************************************************************************************)
METHOD PRIVATE m_ApplyConfig : BOOL
VAR_IN_OUT
	vio_New								: ST_VisuCartesianConfig;
END_VAR
m_ApplyConfig := Tc2_System.MEMCMP(ADR(vio_New), ADR(vo_Visu.stConfig), SIZEOF(vio_New)) <> 0;
IF m_ApplyConfig THEN
	vo_Visu.stConfig := vio_New;
	m_NotifyConfigChanged();
END_IF
END_METHOD

(****************************************************************************************************<br>
© Syntegon Group.<br>
All rights reserved, also regarding any disposal, exploitation, reproduction, editing, distribution,<br>
as well as in the event of applications for industrial property rights.<br>
*****************************************************************************************************<br>
DESCRIPTION:<br>
Manifest type: Cartesian robot.<br>
****************************************************************************************************)
METHOD PROTECTED m_ComponentType : E_VisuComponentType
m_ComponentType := E_VisuComponentType.CARTESIAN;
END_METHOD

(****************************************************************************************************<br>
© Syntegon Group.<br>
All rights reserved, also regarding any disposal, exploitation, reproduction, editing, distribution,<br>
as well as in the event of applications for industrial property rights.<br>
*****************************************************************************************************<br>
DESCRIPTION:<br>
Sets strokes and rail height; its pose (m_SetPose) is the axis origin X = Y = 0 with Z up. TRUE if anything<br>
changed.<br>
****************************************************************************************************)
METHOD m_Configure : BOOL
VAR_INPUT
	vi_lr_XMin							: LREAL;	// [mm]
	vi_lr_XMax							: LREAL;	// [mm]
	vi_lr_YMin							: LREAL;	// [mm]
	vi_lr_YMax							: LREAL;	// [mm]
	vi_lr_ZMin							: LREAL;	// [mm]
	vi_lr_ZMax							: LREAL;	// [mm]
	vi_lr_RailHeight					: LREAL;	// [mm] top of the rails above the local origin
END_VAR
VAR
	TempNew								: ST_VisuCartesianConfig;
END_VAR
TempNew := vo_Visu.stConfig;
TempNew.fXMin := vi_lr_XMin;
TempNew.fXMax := vi_lr_XMax;
TempNew.fYMin := vi_lr_YMin;
TempNew.fYMax := vi_lr_YMax;
TempNew.fZMin := vi_lr_ZMin;
TempNew.fZMax := vi_lr_ZMax;
TempNew.fRailHeight := vi_lr_RailHeight;
m_Configure := m_ApplyConfig(TempNew);
END_METHOD

(****************************************************************************************************<br>
© Syntegon Group.<br>
All rights reserved, also regarding any disposal, exploitation, reproduction, editing, distribution,<br>
as well as in the event of applications for industrial property rights.<br>
*****************************************************************************************************<br>
DESCRIPTION:<br>
The robot's gripper fingers for _FB_VisuRobot.m_SetFinger and m_ClearFingers.<br>
****************************************************************************************************)
METHOD PROTECTED m_Fingers : BOOL
VAR_OUTPUT
	vo_p_Count							: POINTER TO UINT;
	vo_p_Fingers						: POINTER TO ARRAY[0..VISU_GlobalConst_Param.VISU_un_MAX_FINGERS - 1] OF ST_VisuFinger;
END_VAR
vo_p_Count := ADR(vo_Visu.stConfig.nFingerCount);
vo_p_Fingers := ADR(vo_Visu.stConfig.aFingers);
m_Fingers := TRUE;
END_METHOD

(****************************************************************************************************<br>
© Syntegon Group.<br>
All rights reserved, also regarding any disposal, exploitation, reproduction, editing, distribution,<br>
as well as in the event of applications for industrial property rights.<br>
*****************************************************************************************************<br>
DESCRIPTION:<br>
The robot's limit area and TCP limit area for _FB_VisuRobot.m_SetLimitArea, m_ClearLimitArea,<br>
m_SetTcpLimitArea and m_ClearTcpLimitArea.<br>
****************************************************************************************************)
METHOD PROTECTED m_LimitArea : BOOL
VAR_OUTPUT
	vo_p_LimitArea						: POINTER TO ST_VisuLimitArea;
	vo_p_TcpLimitArea					: POINTER TO ST_VisuLimitArea;
END_VAR
vo_p_LimitArea := ADR(vo_Visu.stConfig.stLimitArea);
vo_p_TcpLimitArea := ADR(vo_Visu.stConfig.stTcpLimitArea);
m_LimitArea := TRUE;
END_METHOD

(****************************************************************************************************<br>
© Syntegon Group.<br>
All rights reserved, also regarding any disposal, exploitation, reproduction, editing, distribution,<br>
as well as in the event of applications for industrial property rights.<br>
*****************************************************************************************************<br>
DESCRIPTION:<br>
The pose in vo_Visu, for m_SetPose.<br>
****************************************************************************************************)
METHOD PROTECTED m_Pose : BOOL
VAR_OUTPUT
	vo_p_Pose							: POINTER TO ST_VisuPose;
END_VAR
vo_p_Pose := ADR(vo_Visu.stConfig.stPose);
m_Pose := TRUE;
END_METHOD

(****************************************************************************************************<br>
© Syntegon Group.<br>
All rights reserved, also regarding any disposal, exploitation, reproduction, editing, distribution,<br>
as well as in the event of applications for industrial property rights.<br>
*****************************************************************************************************<br>
DESCRIPTION:<br>
Reports the axes' actual values and the gripper. Call once per cycle; it also stamps the state with the<br>
cycle's DC time.<br>
****************************************************************************************************)
METHOD m_SetAxes : BOOL
VAR_INPUT
	vi_lr_X								: LREAL;	// [mm]
	vi_lr_Y								: LREAL;	// [mm]
	vi_lr_Z								: LREAL;	// [mm]
	vi_b_GripperActive					: BOOL;	// used only when no fingers are configured, else FALSE
END_VAR
vo_Visu.stState.fX := vi_lr_X;
vo_Visu.stState.fY := vi_lr_Y;
vo_Visu.stState.fZ := vi_lr_Z;
vo_Visu.stState.bGripperActive := vi_b_GripperActive;
vo_Visu.stState.nTimestamp := m_DcTime();
m_SetAxes := TRUE;
END_METHOD

(****************************************************************************************************<br>
© Syntegon Group.<br>
All rights reserved, also regarding any disposal, exploitation, reproduction, editing, distribution,<br>
as well as in the event of applications for industrial property rights.<br>
*****************************************************************************************************<br>
DESCRIPTION:<br>
Sets or clears the fault of the robot: drawn red with the message while active. The fault stays until it<br>
is cleared with m_SetFault(vi_b_Active := FALSE, vi_str_Message := ''). TRUE.<br>
****************************************************************************************************)
METHOD m_SetFault : BOOL
VAR_INPUT
	vi_b_Active							: BOOL;	// TRUE: fault active
	vi_str_Message						: STRING(80);	// shown to the operator; empty shows 'Fault'
END_VAR
vo_Visu.stState.stFault.bActive := vi_b_Active;
vo_Visu.stState.stFault.sMessage := vi_str_Message;
m_SetFault := TRUE;
END_METHOD

(****************************************************************************************************<br>
© Syntegon Group.<br>
All rights reserved, also regarding any disposal, exploitation, reproduction, editing, distribution,<br>
as well as in the event of applications for industrial property rights.<br>
*****************************************************************************************************<br>
DESCRIPTION:<br>
Reports finger vi_un_Finger (1-based): the pose of its frame (centre of its top face), absolute in the MCS,<br>
and whether it grips. Call once per cycle per configured finger. A finger never reported here is drawn at its<br>
offset on the flange (m_SetFingerOffset, ADR 0018).<br>
*****************************************************************************************************<br>
OUTPUT VALUES:<br>
FALSE outside 1..VISU_GlobalConst_Param.VISU_un_MAX_FINGERS.<br>
****************************************************************************************************)
METHOD m_SetFingerState : BOOL
VAR_INPUT
	vi_un_Finger						: UINT;	// [-] 1-based
	vi_Pose								: ST_VisuPose;	// MCS
	vi_b_Active							: BOOL;	// TRUE while the finger grips
END_VAR
m_SetFingerState := vi_un_Finger > 0 AND vi_un_Finger <= VISU_GlobalConst_Param.VISU_un_MAX_FINGERS;
IF m_SetFingerState THEN
	vo_Visu.stState.aFingerStates[vi_un_Finger - 1].stPose := vi_Pose;
	vo_Visu.stState.aFingerStates[vi_un_Finger - 1].bActive := vi_b_Active;
	vo_Visu.stState.aFingerStates[vi_un_Finger - 1].bPoseReported := TRUE;
END_IF
END_METHOD

(****************************************************************************************************<br>
© Syntegon Group.<br>
All rights reserved, also regarding any disposal, exploitation, reproduction, editing, distribution,<br>
as well as in the event of applications for industrial property rights.<br>
*****************************************************************************************************<br>
DESCRIPTION:<br>
Sets which axes the robot has. XYZ (default): rails, bridge, carriage and column. XZ: no Y axis, a fixed beam<br>
along the local X at the rail height; the Y stroke and m_SetAxes vi_lr_Y are ignored. XY: no Z axis, the column<br>
has a fixed length and the flange stays at vi_lr_ZMin; vi_lr_ZMax and m_SetAxes vi_lr_Z are ignored.<br>
TRUE if anything changed.<br>
****************************************************************************************************)
METHOD m_SetKinematics : BOOL
VAR_INPUT
	vi_e_Axes							: E_VisuCartesianAxes;	// axes of the robot
END_VAR
VAR
	TempNew								: ST_VisuCartesianConfig;
END_VAR
TempNew := vo_Visu.stConfig;
TempNew.eAxes := vi_e_Axes;
m_SetKinematics := m_ApplyConfig(TempNew);
END_METHOD

(****************************************************************************************************<br>
© Syntegon Group.<br>
All rights reserved, also regarding any disposal, exploitation, reproduction, editing, distribution,<br>
as well as in the event of applications for industrial property rights.<br>
*****************************************************************************************************<br>
DESCRIPTION:<br>
Moves the robot's shown coordinate system (origin triad, local measuring coordinates) away from axis zero<br>
(stPose), in the robot's local frame. Geometry and axis values stay relative to stPose. TRUE if anything changed.<br>
****************************************************************************************************)
METHOD m_SetOriginShift : BOOL
VAR_INPUT
	vi_lr_X								: LREAL;	// [mm] along the robot's local X
	vi_lr_Y								: LREAL;	// [mm] along the robot's local Y, 0 = none
	vi_lr_Z								: LREAL;	// [mm] along the robot's local Z, 0 = none
END_VAR
VAR
	TempNew								: ST_VisuCartesianConfig;
END_VAR
TempNew := vo_Visu.stConfig;
TempNew.stOriginShift.fX := vi_lr_X;
TempNew.stOriginShift.fY := vi_lr_Y;
TempNew.stOriginShift.fZ := vi_lr_Z;
m_SetOriginShift := m_ApplyConfig(TempNew);
END_METHOD

(****************************************************************************************************<br>
© Syntegon Group.<br>
All rights reserved, also regarding any disposal, exploitation, reproduction, editing, distribution,<br>
as well as in the event of applications for industrial property rights.<br>
*****************************************************************************************************<br>
DESCRIPTION:<br>
The robot's zones for _FB_VisuZoneComponent.m_SetZone and m_ClearZones.<br>
****************************************************************************************************)
METHOD PROTECTED m_Zones : BOOL
VAR_OUTPUT
	vo_p_Count							: POINTER TO UINT;
	vo_p_Zones							: POINTER TO ARRAY[0..VISU_GlobalConst_Param.VISU_un_MAX_ZONES - 1] OF ST_VisuZone;
END_VAR
vo_p_Count := ADR(vo_Visu.stConfig.nZoneCount);
vo_p_Zones := ADR(vo_Visu.stConfig.aZones);
m_Zones := TRUE;
END_METHOD

END_FUNCTION_BLOCK

// POUs/_FB_VisuMachine
(****************************************************************************************************<br>
© Syntegon Group.<br>
All rights reserved, also regarding any disposal, exploitation, reproduction, editing, distribution,<br>
as well as in the event of applications for industrial property rights.<br>
*****************************************************************************************************<br>
DESCRIPTION:<br>
The machine as its application reports it (protocol 22, ADR 0021): run state, simulation mode and machine<br>
messages, written to the machine entry GVL_Visu.stMachine next to the manifest. Not a component: it has no<br>
manifest entry. The application calls m_Register and the other methods every cycle; a machine message is set by<br>
its level (m_SetMessage), like a component's fault.<br>
*****************************************************************************************************<br>
VERSION         ¦ DATE       ¦ NAME      ¦ CHANGE<br>
Syn_Visu 9.7.0  ¦ 2026-11-13 ¦ J.Willner ¦ Created: run state, simulation mode, machine messages (protocol 22)<br>
****************************************************************************************************)
FUNCTION_BLOCK _FB_VisuMachine
VAR
	RefMachine							: REFERENCE TO ST_VisuMachine;	// set by m_Register
END_VAR

(****************************************************************************************************<br>
© Syntegon Group.<br>
All rights reserved, also regarding any disposal, exploitation, reproduction, editing, distribution,<br>
as well as in the event of applications for industrial property rights.<br>
*****************************************************************************************************<br>
DESCRIPTION:<br>
Distributed-clock time of the calling task's current cycle in ns since 2000-01-01; 0 if unknown.<br>
****************************************************************************************************)
METHOD PRIVATE m_DcTime : ULINT
VAR
	dn_TempTaskIndex					: DINT;
END_VAR
dn_TempTaskIndex := Tc2_System.GETCURTASKINDEXEX();
IF dn_TempTaskIndex > 0 THEN
	m_DcTime := LINT_TO_ULINT(TwinCAT_SystemInfoVarList._TaskInfo[dn_TempTaskIndex].DcTaskTime);
ELSE
	m_DcTime := 0;
END_IF
END_METHOD

(****************************************************************************************************<br>
© Syntegon Group.<br>
All rights reserved, also regarding any disposal, exploitation, reproduction, editing, distribution,<br>
as well as in the event of applications for industrial property rights.<br>
*****************************************************************************************************<br>
DESCRIPTION:<br>
Connects this block to the application's machine entry, GVL_Visu.stMachine. Call it every cycle before the other<br>
methods, which also keeps the reference valid after an online change.<br>
*****************************************************************************************************<br>
OUTPUT VALUES:<br>
Always TRUE.<br>
****************************************************************************************************)
METHOD m_Register : BOOL
VAR_IN_OUT
	vio_Machine							: ST_VisuMachine;	// GVL_Visu.stMachine of the application
END_VAR
RefMachine REF= vio_Machine;
m_Register := TRUE;
END_METHOD

